FUNCTION_BLOCK FB_BECKHOFF_AxisController
(*

The function block used to control axis.

Constructor: 		Patryk Panylo
Company:		E. Riexinger GmbH
Date:			23.04.2015
Version:			1.00

Date:			Revision:		Who:				Comment
dd.mm.yyyy		x.xx			Initials			comment

*)
VAR_INPUT
	(* Input variables / Eingang Variablen *)
	bEnable						:BOOL;						(* Signal FB enable *)
	etMachineMode				:ET_MachineMode;			(* Machine mode *)
	etMachineState				:ET_MachineState;			(* Machine state *)
	bNoEStop					:BOOL;						(* No ermergency Stop / Keine Notaus *)
	bRegulatorOn				:BOOL;						(* Enable the power stage *)
	bReset						:BOOL;						(* Signal reset *)
	bCMDInterrupt				:BOOL;						(* Signal interrupt *)
	bTerminalOK					:BOOL;						(* Terminal Ok *)
	bExeReset					:BOOL;						(* Execute auto reset *)
	bExeSetPos					:BOOL;						(* Execute set position *)
	lrSetPosition				:LREAL;						(* Position value to which the axis position is to be set. *)
	bExeGearIn					:BOOL;						(* Execute gear in *)
	bExeGearOut					:BOOL;						(* Execute gear out *)
	dnRatioNumerator			:DINT;						(* Gear ratio numerator. Alternatively, the gear ratio can be specified in the numerator as a floating comma value, if the denominator is 1. *)
	udnRatioDenominator			:UDINT;						(* Gear ratio denominator *)
	lrOverride					:LREAL;						(* Override 100% percent *)
	bWithAbsoluteEncoder		:BOOL; 						(* Encoder is an absolute one / Absolutwertgeber *)
	bPosLagMonitoringEn			:BOOL;						(* Enable position lag monitoring *)
	lrPositionBias				:LREAL;						(* Position bias *)
	bHWSignalLimitMax			:BOOL;						(* Signal position limit switch maximum *)
	bHWSignalLimitMin			:BOOL;						(* Signal position limit switch minimum *)
	lrSoftLimitMax				:LREAL; 					(* Position limit switch maximum *)
	lrSoftLimitMin				:LREAL; 					(* Position limit switch minimum *)
	lrAcceleration				:LREAL;						(* Value of the acceleration (always positive) *)
	lrDeceleration				:LREAL;						(* Value of deceleration (always positive) *)
	lrJerk						:LREAL;						(* Value of jerk (always positive) *)
	lrActTemp					:LREAL;						(* Current temperatur *)
	tAdsTimeOut 				:TIME := T#2S;				(* Timout for ads commands *)
END_VAR
VAR_OUTPUT
	(* Output variables / Ausgang Variablen *)
	bStatus						:BOOL;						(* Feedback *)
	bStatusDelay				:BOOL;						(* Feedback delay *)
	bReseted					:BOOL;						(* Reset completed *)
	bError						:BOOL;						(* Controller error *)
	bErrorInit					:BOOL;						(* Controller initialization error *)
	udnErrorNo					:UDINT;						(* Error number *)
	lrActPos					:LREAL;						(* Actual position *)
	lrSetPos					:LREAL;						(* Set position *)
	lrActAbsPos					:LREAL;						(* Actual absolut position *)
	lrActVelo					:LREAL;						(* Actual velocity *)
	bNotMoving					:BOOL;						(* Status of moving *)
	bReferenced					:BOOL;						(* Referenced *)
	bCoupled					:BOOL;						(* Coupled *)
	lrVeloLimitMax				:LREAL;						(* Velocity limit maximum *)
	lrAccLimitMax				:LREAL;						(* Acceleration limit maximum *)
	lrDecLimitMax				:LREAL;						(* Deceleration limit maximum *)
	lrJerkLimitMax				:LREAL;						(* Jerk limit maximum *)
	bHardLimitMaxExceeded		:BOOL;						(* Position limit switch maximum is exceeded *)
	bHardLimitMinExceeded		:BOOL;						(* Position limit switch minimum is exceeded *)
	bSoftLimitMaxExceeded		:BOOL;						(* Position limit switch maximum is exceeded *)
	bSoftLimitMinExceeded		:BOOL;						(* Position limit switch minimum is exceeded *)
END_VAR
VAR_IN_OUT
	Axis						:AXIS_REF;					(* The AXIS_REF data type  is an interface between the PLC and the NC and contains axis information *)
	MasterAxis					:AXIS_REF;					(* The AXIS_REF data type  is an interface between the PLC and the NC and contains axis information *)
END_VAR
VAR
	(* Enummerations *)

	(* Variables *)
	etAxisGetLimits				:ET_BECKHOFF_AxisGetLimits;
	bGetLimitsExe				:BOOL;						(* Progam execute *)
	bGetLimitsDone 				:BOOL;                      (* Program done *)
	bGetLimitsBusy 				:BOOL;                      (* Program busy *)
	bGetLimitsError 			:BOOL;                      (* Program error *)
	bGetLimitsInitDone 			:BOOL;                      (* Program initialization done *)
	udnGetLimitsErrorNo 		:UDINT;                     (* Error number *)
	unGetValueWatchdog			:UINT;

	etAxisSetLimits				:ET_BECKHOFF_AxisSetLimits;
	bSetLimitsExe				:BOOL;						(* Progam execute *)
	bSetLimitsDone 				:BOOL;                      (* Program done *)
	bSetLimitsBusy 				:BOOL;                      (* Program busy *)
	bSetLimitsError 			:BOOL;                      (* Program error *)
	bSetLimitsInitDone 			:BOOL;                      (* Program initialization done *)
	bSetLimitsInitError 		:BOOL;                      (* Program initialization error *)
	udnSetLimitsErrorNo 		:UDINT;                     (* Error number *)
	unSetValueWatchdog			:UINT;

	tStatusDelay				:TIME := T#1S;				(* Status delay time *)
	tRegulatorOffDelay			:TIME := T#50MS;			(* Regulator off delay time *)

	dwReferenceSystem			:DWORD;						(* Reference system: 0 - INC, 1 - ABS, 2 - ABS MODULO *)
	lrPositionBiasCache			:LREAL;						(* Position bias *)
	lrSoftLimitMaxCache			:LREAL; 					(* Position limit switch maximum *)
	lrSoftLimitMinCache			:LREAL; 					(* Position limit switch minimum *)

	tonFirstInit				:TON;						(* First initialization *)
	bFirstTime					:BOOL;

	(* References *)

	(* Interfaces *)

	(* Instances *)
	fbMcPower					:MC_Power;					(* The function block is used to enable for an axis *)
	rtNoEStop					:R_TRIG;
	tofRegulatorOn				:TOF;						(* Delay controller disable *)
	tonStatusDelay				:TON;						(* Delay controller enabled status *)
	fbMcReset					:MC_Reset;					(* An axis reset is carried out with the function block *)
	fbMcSetPosition				:MC_SetPosition;			(* Sets the current axis position to a parameterisable value. *)
	fbMcGearIn					:MC_GearInDyn;				(* The function block is used to couples a slave axis to a master axis using a floating point gear ratio. *)
	fbMcGearOut					:MC_GearOut;				(* The function block  is used to decoupling the slave from the master axis.  *)
	fbMcReadParameter 			:MC_ReadParameter;			(* The function block is used to read an axis parameter. *)
	fbMcWriteParameter 			:MC_WriteParameter;			(* The function block is used to write an axis parameter. *)
	fbMcWriteBoolParameter 		:MC_WriteBoolParameter;		(* The function block is used to write bool value an axis parameter. *)
	fbAdsWrite					:ADSWRITE;					(* The function block permits execution of an ADS write command, for the transfer of data to an ADS device. *)
	fbAdsRead					:ADSREAD;					(* The function block permits execution of an ADS read command, for the transfer of data to an ADS device. *)
	tofRepeateSetLimitsInit		:TOF;
	tofRepeateGetLimitsInit		:TOF;
	tonCoupled					:TON;
END_VAR
VAR CONSTANT
	dwIdxGrMainPara				:DWORD := 16#00004000;		(* Index group for main parameters of axis *)
	dwIdxGrNCEncPara			:DWORD := 16#00005000;		(* Index group for nc-encoder parameters of axis *)
	dwIdxGrNCCtrlPara			:DWORD := 16#00006000;		(* Index group for nc-controller parameters of axis *)
	dwIdxGrNCDrivePara			:DWORD := 16#00007000;		(* Index group for nc-drive parameters of axis *)
	
	tFirstInit					:TIME := T#2S;				(* First initialization *)
	tRepeateInit				:TIME := T#1S;				(* Repeate initialization *)
	
	unWatchdogMax				:UINT := 150;
END_VAR

IF NOT bEnable							(* Signal FB enable *)
THEN
	bStatus := FALSE;						(* Feedback *)
	bStatusDelay := FALSE;				(* Feedback *)
	bError := FALSE;						(* Controller error *)
	udnErrorNo := 0;						(* Error number *)

	bFirstTime := FALSE;
	RETURN;
END_IF

IF NOT bFirstTime
THEN
	tonFirstInit(IN := FALSE);					(* Program execute *)
	bGetLimitsDone := FALSE;                                	(* Program done *)
	bGetLimitsBusy := FALSE;                                 	(* Program not busy *)
	bGetLimitsError := FALSE;                                 	(* Program not error *)
	bGetLimitsInitDone := FALSE;				(* Program initialization done *)
	udnGetLimitsErrorNo := 0;                                 		(* Error number *)
	unGetValueWatchdog := 0;

	etAxisGetLimits := ET_BECKHOFF_AxisGetLimits.eWaitExecute;       			(* Next step *)

	bSetLimitsExe := FALSE;					(* Program execute *)
	bSetLimitsDone := FALSE;                                	(* Program done *)
	bSetLimitsBusy := FALSE;                                 	(* Program not busy *)
	bSetLimitsError := FALSE;                                	 	(* Program not error *)
	bSetLimitsInitDone := FALSE;                            	(* Program initialization done *)
	bSetLimitsInitError := FALSE;				(* Program initialization error *)
	udnSetLimitsErrorNo := 0;                                 		(* Error number *)
	unSetValueWatchdog := 0;
	
	etAxisSetLimits := ET_BECKHOFF_AxisSetLimits.eWaitExecute;       			(* Next step *)

	(* Actual position *)
	lrActAbsPos := Axis.NcToPlc.ActPos;
	lrActAbsPos := F_LRealRound(lrReal := lrActAbsPos, usiPrecision := 3);

	bFirstTime := TRUE;
END_IF;

A_MCPower();
A_MCReset();
A_MCSetPosition();
A_MCGearCoupling();
A_Utility();
A_GetLimits();
A_SetLimits();
A_Error();

(* Actual position *)
lrActPos := Axis.NcToPlc.ActPos;
lrActPos := F_LRealRound(lrReal := lrActPos, usiPrecision := 2);

(* Set position *)
lrSetPos := Axis.NcToPlc.SetPos;
lrSetPos := F_LRealRound(lrReal := lrSetPos, usiPrecision := 2);

(* Actual velocity *)
lrActVelo := Axis.NcToPlc.ActVelo;
lrActVelo := F_LRealRound(lrReal := lrActVelo, usiPrecision := 2);

(* Current engine torque *)
(*nActEngineTorque := Axis.stNcToPlc.stCommandPositioning.nActEngineTorque;*)

(* Reference signal *)
bReferenced := Axis.NcToPlc.StateDWord.1;                               (* In Reference *)


(* Status not moving *)
bNotMoving := Axis.NcToPlc.StateDWord.2;

(* Status coupling *)
tonCoupled(
	IN := Axis.NcToPlc.CoupleState = 2
		  OR Axis.NcToPlc.CoupleState = 3,
	PT := T#200MS
);
bCoupled := tonCoupled.Q;

ACTION A_Error:

bError := fbMcPower.Error
		OR fbMcReset.Error
	  	OR fbMcSetPosition.Error
		OR fbMcGearIn.Error
		OR fbMcGearOut.Error
		OR Axis.NcToPlc.StateDWord.31
		OR MasterAxis.NcToPlc.StateDWord.31;

bErrorInit := bGetLimitsError
		      OR bSetLimitsError;
END_ACTION

ACTION A_GetLimits:

(* Status hardware limit switch *)
bHardLimitMaxExceeded := bHWSignalLimitMax;						(* Position limit switch maximum is exceeded *)
bHardLimitMinExceeded := bHWSignalLimitMin;						(* Position limit switch minimum is exceeded *)

(* Status software limit switch *)
bSoftLimitMaxExceeded := Axis.NcToPlc.StateDWord.27 AND lrSoftLimitMax <> lrSoftLimitMin;	(* Position limit switch maximum is exceeded *)
bSoftLimitMinExceeded := Axis.NcToPlc.StateDWord.26 AND lrSoftLimitMax <> lrSoftLimitMin;		(* Position limit switch minimum is exceeded *)

(* Get limits execute *)
tofRepeateGetLimitsInit(
	IN := bGetLimitsError,
	PT := tRepeateInit
);

tonFirstInit(
	IN:= bTerminalOK
		 AND NOT bGetLimitsInitDone,
	PT := tFirstInit
);

bGetLimitsExe := (tonFirstInit.Q
				  OR bGetLimitsInitDone)
				  AND NOT tofRepeateGetLimitsInit.Q;

(* Get axis limits *)
CASE etAxisGetLimits OF

	ET_BECKHOFF_AxisGetLimits.eWaitExecute:
		IF bGetLimitsExe
		   AND bTerminalOK
		THEN
			unGetValueWatchdog := 0;
			bGetLimitsDone := FALSE;                                	(* Program done *)
			bGetLimitsBusy := FALSE;                                 	(* Program not busy *)
			bGetLimitsError := FALSE;                                 	(* Program not error *)
			udnGetLimitsErrorNo := 0;                                 	(* Error number *)

			fbMcReadParameter(
				Enable:= FALSE,
				ReadMode := READMODE_ONCE,
				Axis := Axis
			);

			fbAdsRead(
				NETID := '',
				READ := FALSE,
				TMOUT := tAdsTimeOut
			);
			
			etAxisGetLimits := ET_BECKHOFF_AxisGetLimits.eReadVeloMax;         		(* Next step *)
		END_IF

	ET_BECKHOFF_AxisGetLimits.eReadVeloMax:
		fbMcReadParameter.Enable := TRUE;
		fbMcReadParameter.ParameterNumber:= MaxVelocityAppl;

		unGetValueWatchdog := unGetValueWatchdog + 1;
		
		IF fbMcReadParameter.Busy
		THEN
			etAxisGetLimits := ET_BECKHOFF_AxisGetLimits.eWfReadVeloMax;         		(* Next step *)

		ELSIF fbMcReadParameter.Error
		THEN
			fbMcReadParameter(
				Enable:= FALSE,
				Axis := Axis
			);

			udnGetLimitsErrorNo := 1;                                 	(* Error number *)
			
			etAxisGetLimits := ET_BECKHOFF_AxisGetLimits.eError;         		(* Next step *)

		END_IF

	ET_BECKHOFF_AxisGetLimits.eWfReadVeloMax:
		IF NOT fbMcReadParameter.Busy
		     AND NOT fbMcReadParameter.Error
		THEN
			fbMcReadParameter(
				Enable:= FALSE,
				Axis := Axis
			);

			lrVeloLimitMax := fbMcReadParameter.Value;

			unGetValueWatchdog := 0;
			
			etAxisGetLimits := ET_BECKHOFF_AxisGetLimits.eReadAccMax;         		(* Next step *)

		ELSIF fbMcReadParameter.Error
		THEN
			fbMcReadParameter(
				Enable:= FALSE,
				Axis := Axis
			);

			udnGetLimitsErrorNo := 2;                                 	(* Error number *)
			
			etAxisGetLimits := ET_BECKHOFF_AxisGetLimits.eError;         		(* Next step *)

		END_IF

	ET_BECKHOFF_AxisGetLimits.eReadAccMax:
		fbMcReadParameter.Enable := TRUE;
		fbMcReadParameter.ParameterNumber:= MaxAccelerationAppl;

		unGetValueWatchdog := unGetValueWatchdog + 1;
		
		IF fbMcReadParameter.Busy
		THEN
			etAxisGetLimits := ET_BECKHOFF_AxisGetLimits.eWfReadAccMax;         		(* Next step *)

		ELSIF fbMcReadParameter.Error
		THEN
			fbMcReadParameter(
				Enable:= FALSE,
				Axis := Axis
			);

			udnGetLimitsErrorNo := 3;                                 	(* Error number *)
			
			etAxisGetLimits := ET_BECKHOFF_AxisGetLimits.eError;         		(* Next step *)

		END_IF

	ET_BECKHOFF_AxisGetLimits.eWfReadAccMax:
		IF NOT fbMcReadParameter.Busy
		     AND NOT fbMcReadParameter.Error
		THEN
			fbMcReadParameter(
				Enable:= FALSE,
				Axis := Axis
			);

			lrAccLimitMax := fbMcReadParameter.Value;

			unGetValueWatchdog := 0;
			
			etAxisGetLimits := ET_BECKHOFF_AxisGetLimits.eReadDecMax;         		(* Next step *)

		ELSIF fbMcReadParameter.Error
		THEN
			fbMcReadParameter(
				Enable:= FALSE,
				Axis := Axis
			);

			udnGetLimitsErrorNo := 4;                                 	(* Error number *)
			
			etAxisGetLimits := ET_BECKHOFF_AxisGetLimits.eError;         		(* Next step *)

		END_IF

	ET_BECKHOFF_AxisGetLimits.eReadDecMax:
		fbMcReadParameter.Enable := TRUE;
		fbMcReadParameter.ParameterNumber:= MaxDecelerationAppl;

		unGetValueWatchdog := unGetValueWatchdog + 1;
		
		IF fbMcReadParameter.Busy
		THEN
			etAxisGetLimits := ET_BECKHOFF_AxisGetLimits.eWfReadDecMax;         		(* Next step *)

		ELSIF fbMcReadParameter.Error
		THEN
			fbMcReadParameter(
				Enable:= FALSE,
				Axis := Axis
			);

			udnGetLimitsErrorNo := 5;                                 	(* Error number *)
			
			etAxisGetLimits := ET_BECKHOFF_AxisGetLimits.eError;         		(* Next step *)

		END_IF

	ET_BECKHOFF_AxisGetLimits.eWfReadDecMax:
		IF NOT fbMcReadParameter.Busy
		     AND NOT fbMcReadParameter.Error
		THEN
			fbMcReadParameter(
				Enable:= FALSE,
				Axis := Axis
			);

			lrDecLimitMax := fbMcReadParameter.Value;

			unGetValueWatchdog := 0;
			
			etAxisGetLimits := ET_BECKHOFF_AxisGetLimits.eReadJerkMax;         		(* Next step *)

		ELSIF fbMcReadParameter.Error
		THEN
			fbMcReadParameter(
				Enable:= FALSE,
				Axis := Axis
			);

			udnGetLimitsErrorNo := 6;                                 	(* Error number *)
			
			etAxisGetLimits := ET_BECKHOFF_AxisGetLimits.eError;         		(* Next step *)

		END_IF

	ET_BECKHOFF_AxisGetLimits.eReadJerkMax:
		fbMcReadParameter.Enable := TRUE;
		fbMcReadParameter.ParameterNumber:= MaxJerkAppl;

		unGetValueWatchdog := unGetValueWatchdog + 1;
		
		IF fbMcReadParameter.Busy
		THEN
			etAxisGetLimits := ET_BECKHOFF_AxisGetLimits.eWfReadJerkMax;         		(* Next step *)

		ELSIF fbMcReadParameter.Error
		THEN
			fbMcReadParameter(
				Enable:= FALSE,
				Axis := Axis
			);

			udnGetLimitsErrorNo := 7;                                 	(* Error number *)
			
			etAxisGetLimits := ET_BECKHOFF_AxisGetLimits.eError;         		(* Next step *)

		END_IF

	ET_BECKHOFF_AxisGetLimits.eWfReadJerkMax:
		IF NOT fbMcReadParameter.Busy
		     AND NOT fbMcReadParameter.Error
		THEN
			fbMcReadParameter(
				Enable:= FALSE,
				Axis := Axis
			);

			lrJerkLimitMax := fbMcReadParameter.Value;

			unGetValueWatchdog := 0;
			
			etAxisGetLimits := ET_BECKHOFF_AxisGetLimits.eReadSoftLimitMax;         		(* Next step *)

		ELSIF fbMcReadParameter.Error
		THEN
			fbMcReadParameter(
				Enable:= FALSE,
				Axis := Axis
			);

			udnGetLimitsErrorNo := 8;                                 	(* Error number *)
			
			etAxisGetLimits := ET_BECKHOFF_AxisGetLimits.eError;         		(* Next step *)

		END_IF

	ET_BECKHOFF_AxisGetLimits.eReadSoftLimitMax:
		fbMcReadParameter.Enable := TRUE;
		fbMcReadParameter.ParameterNumber:= SWLimitPos;

		unGetValueWatchdog := unGetValueWatchdog + 1;
		
		IF fbMcReadParameter.Busy
		THEN
			etAxisGetLimits := ET_BECKHOFF_AxisGetLimits.eWfReadSoftLimitMax;         		(* Next step *)

		ELSIF fbMcReadParameter.Error
		THEN
			fbMcReadParameter(
				Enable:= FALSE,
				Axis := Axis
			);

			udnGetLimitsErrorNo := 9;                                 	(* Error number *)
			
			etAxisGetLimits := ET_BECKHOFF_AxisGetLimits.eError;         		(* Next step *)

		END_IF

	ET_BECKHOFF_AxisGetLimits.eWfReadSoftLimitMax:
		IF NOT fbMcReadParameter.Busy
		     AND NOT fbMcReadParameter.Error
		THEN
			fbMcReadParameter(
				Enable:= FALSE,
				Axis := Axis
			);

			lrSoftLimitMax := fbMcReadParameter.Value;

			unGetValueWatchdog := 0;
			
			etAxisGetLimits := ET_BECKHOFF_AxisGetLimits.eReadSoftLimitMin;         		(* Next step *)

		ELSIF fbMcReadParameter.Error
		THEN
			fbMcReadParameter(
				Enable:= FALSE,
				Axis := Axis
			);

			udnGetLimitsErrorNo := 10;                                 	(* Error number *)
			
			etAxisGetLimits := ET_BECKHOFF_AxisGetLimits.eError;         		(* Next step *)

		END_IF

	ET_BECKHOFF_AxisGetLimits.eReadSoftLimitMin:
		fbMcReadParameter.Enable := TRUE;
		fbMcReadParameter.ParameterNumber:= SWLimitNeg;

		unGetValueWatchdog := unGetValueWatchdog + 1;
		
		IF fbMcReadParameter.Busy
		THEN
			etAxisGetLimits := ET_BECKHOFF_AxisGetLimits.eWfReadSoftLimitMin;         		(* Next step *)

		ELSIF fbMcReadParameter.Error
		THEN
			fbMcReadParameter(
				Enable:= FALSE,
				Axis := Axis
			);

			udnGetLimitsErrorNo := 11;                                 	(* Error number *)
			
			etAxisGetLimits := ET_BECKHOFF_AxisGetLimits.eError;         		(* Next step *)

		END_IF

	ET_BECKHOFF_AxisGetLimits.eWfReadSoftLimitMin:
		IF NOT fbMcReadParameter.Busy
		     AND NOT fbMcReadParameter.Error
		THEN
			fbMcReadParameter(
				Enable:= FALSE,
				Axis := Axis
			);

			lrSoftLimitMin := fbMcReadParameter.Value;

			unGetValueWatchdog := 0;
			
			etAxisGetLimits := ET_BECKHOFF_AxisGetLimits.eDone;         		(* Next step *)

		ELSIF fbMcReadParameter.Error
		THEN
			fbMcReadParameter(
				Enable:= FALSE,
				Axis := Axis
			);

			udnGetLimitsErrorNo := 12;                                 	(* Error number *)
			
			etAxisGetLimits := ET_BECKHOFF_AxisGetLimits.eError;         		(* Next step *)

		END_IF
	
	ET_BECKHOFF_AxisGetLimits.eDone:
		bGetLimitsDone := TRUE;                                     		(* Program done, in position *)
		bGetLimitsBusy := FALSE;                                     		(* Program not busy *)
		bGetLimitsInitDone := TRUE;                             		(* Program initialization done *)

		etAxisGetLimits := ET_BECKHOFF_AxisGetLimits.eNoExecute;            	(* Next step *)

	ET_BECKHOFF_AxisGetLimits.eError:
		bGetLimitsDone := FALSE;                                     		(* Program done, in position *)
		bGetLimitsError := TRUE;                                     		(* Program error *)
		bGetLimitsBusy := FALSE;                                     		(* Program not busy *)
		bGetLimitsInitDone := FALSE;                             		(* Program initialization done *)

		etAxisGetLimits := ET_BECKHOFF_AxisGetLimits.eNoExecute;           	(* Next step *)

	ET_BECKHOFF_AxisGetLimits.eNoExecute:
		IF NOT bGetLimitsExe
		THEN
			bGetLimitsDone := FALSE;                                     		(* Program done, in position *)
			bGetLimitsError := FALSE;                                     		(* Program error *)
			bGetLimitsBusy := FALSE;                                     		(* Program not busy *)

			etAxisGetLimits := ET_BECKHOFF_AxisGetLimits.eWaitExecute;       (* Next step *)
		END_IF

END_CASE;

fbMcReadParameter(
	ReadMode := READMODE_ONCE,
	Axis := Axis
);
END_ACTION

ACTION A_MCGearCoupling:

(* The function block MC_GearInDyn couples a slave axis to a master axis using a floating point gear ratio. The gear ratio can be dynamically modified every PLC cycle as long as the Execute input is TRUE *)
IF udnRatioDenominator = 0
THEN
	fbMCGearIn.GearRatio := 0;
ELSE
	fbMCGearIn.GearRatio:= dnRatioNumerator / udnRatioDenominator;
END_IF


IF NOT bCMDInterrupt
THEN

	(* The function block MC_GearIn used to coupling with ratio between the velocity of the slave and master axis  *)
	fbMCGearIn(
		Enable := bExeGearIn,
		Acceleration := lrAcceleration,
		Deceleration := lrDeceleration,
		Jerk := lrJerk,
		Options := ,
		Master := MasterAxis,
		Slave := Axis
	);
	
	(* The function block MC_GearOut used to decoupling the Slave from the Master axis.  *)
	fbMCGearOut(
		Execute := bExeGearOut,
		Slave := Axis,
	);

	(* Weiter für die GearIn und GearOut entwickeln*)
	(*Axis.bCmdInterrupted := FALSE;*)

ELSE
	(* The function block MC_GearIn used to coupling with ratio between the velocity of the slave and master axis  *)
	fbMCGearIn(
		Enable := FALSE,
		Master := MasterAxis,
		Slave := Axis
	);

	(* The function block MC_GearOut used to decoupling the Slave from the Master axis.  *)
	fbMCGearOut(
		Execute := FALSE,
		Slave := Axis
	);

	(*Axis.bCmdInterrupted := TRUE;*)
END_IF
END_ACTION

ACTION A_MCPower:

tofRegulatorOn(
	IN := bRegulatorOn,
	PT := tRegulatorOffDelay
);

fbMCPower(
	Enable := tofRegulatorOn.Q
			OR Axis.Status.Moving,
	Enable_Positive := (bRegulatorOn
					AND NOT bHWSignalLimitMax)                          			(* HW limit switch maximum *)
					OR Axis.NcToPlc.HomingState <> 0,
	Enable_Negative := (bRegulatorOn
					   AND NOT bHWSignalLimitMin)                         			(* HW Limit switch minimum *)
					   OR Axis.NcToPlc.HomingState <> 0,
	Override := LIMIT(0.0, lrOverride, 100.0),
	Axis := Axis,
	Status => bStatus,
);

tonStatusDelay(
	IN := fbMCPower.Status,
	PT := SEL(etMachineMode = ET_MachineMode_eManual, tStatusDelay, t#0s),
	Q => bStatusDelay
);
END_ACTION

ACTION A_MCReset:

rtNoEStop(CLK := bNoEStop);

fbMCReset(
	Execute := rtNoEStop.Q
			   OR (bReset
			   		AND Axis.NcToPlc.StateDWord.31)
			   OR bExeReset,
	Axis := Axis,
	Done => bReseted
 );
END_ACTION

ACTION A_MCSetPosition:

fbMCSetPosition(
	Execute := bExeSetPos,
	Position := SEL(lrSoftLimitMin <> lrSoftLimitMax, lrSetPosition, LIMIT(lrSoftLimitMin, lrSetPosition, lrSoftLimitMax)),
	Mode := FALSE,
	Options := ,
	Axis := Axis
);
END_ACTION

ACTION A_SetLimits:

(* Set limits execute *)
tofRepeateSetLimitsInit(
	IN := bSetLimitsError,
	PT := tRepeateInit
);

bSetLimitsExe := SEL(
						bSetLimitsInitDone,
						NOT bSetLimitsInitError,
						NOT bSetLimitsInitError
						AND (lrPositionBias <> lrPositionBiasCache
							   OR lrSoftLimitMaxCache <> lrSoftLimitMax
							   OR lrSoftLimitMinCache <> lrSoftLimitMin)
					);

(* Set axis limits *)
CASE etAxisSetLimits OF

	ET_BECKHOFF_AxisSetLimits.eWaitExecute:
		IF bSetLimitsExe
		   AND bTerminalOK
		   AND bNotMoving
		   AND bGetLimitsDone
		THEN
			unSetValueWatchdog := 0;
			bSetLimitsDone := FALSE;                                	(* Program done *)
			bSetLimitsBusy := FALSE;                                 	(* Program not busy *)
			bSetLimitsError := FALSE;                                	 	(* Program not error *)
			udnSetLimitsErrorNo := 0;                                 		(* Error number *)

			fbMcWriteParameter(
				Execute := FALSE,
				Axis := Axis
			);
	
			fbMcWriteBoolParameter(
				Execute := FALSE,
				Axis := Axis
			);
	
			fbAdsWrite(
				NETID := '',
				WRITE := FALSE,
				TMOUT := tAdsTimeOut
			 );

			etAxisSetLimits := ET_BECKHOFF_AxisSetLimits.eSetReferenceSystem;         		(* Next step *)

		END_IF;

	ET_BECKHOFF_AxisSetLimits.eSetReferenceSystem:
		dwReferenceSystem := BOOL_TO_DWORD(bWithAbsoluteEncoder);

		fbAdsWrite.PORT := 501;
		fbAdsWrite.WRITE := TRUE;
		fbAdsWrite.IDXGRP := dwIdxGrNCEncPara + Axis.NcToPlc.AxisId;
		fbAdsWrite.IDXOFFS := 16#00000019;
		fbAdsWrite.LEN := SIZEOF(dwReferenceSystem);
		fbAdsWrite.SRCADDR := ADR(dwReferenceSystem);

		unSetValueWatchdog := unSetValueWatchdog + 1;
		
		IF fbAdsWrite.Busy
		THEN
			etAxisSetLimits := ET_BECKHOFF_AxisSetLimits.eWfSetReferenceSystem;         		(* Next step *)

		ELSIF fbAdsWrite.ERR
		THEN
			fbAdsWrite(
				WRITE := FALSE,
			);

			udnSetLimitsErrorNo := 1;                                 		(* Error number *)
			
			etAxisSetLimits := ET_BECKHOFF_AxisSetLimits.eError;         		(* Next step *)

		END_IF

	ET_BECKHOFF_AxisSetLimits.eWfSetReferenceSystem:
		IF NOT fbAdsWrite.Busy
		     AND NOT fbAdsWrite.ERR
		THEN
			fbAdsWrite(
				WRITE := FALSE,
			);

			unSetValueWatchdog := 0;
			
			etAxisSetLimits := ET_BECKHOFF_AxisSetLimits.eSetPositionBias;         		(* Next step *)

		ELSIF fbAdsWrite.ERR
		THEN
			fbAdsWrite(
				WRITE := FALSE,
			);

			udnSetLimitsErrorNo := 2;                                 		(* Error number *)
			
			etAxisSetLimits := ET_BECKHOFF_AxisSetLimits.eError;         		(* Next step *)

		END_IF

	ET_BECKHOFF_AxisSetLimits.eSetPositionBias:
		IF bWithAbsoluteEncoder
		THEN
			lrPositionBiasCache := lrPositionBias;

			fbAdsWrite.PORT := 501;
			fbAdsWrite.WRITE := TRUE;
			fbAdsWrite.IDXGRP := dwIdxGrNCEncPara + Axis.NcToPlc.AxisId;
			fbAdsWrite.IDXOFFS := 16#00000007;
			fbAdsWrite.LEN := SIZEOF(lrPositionBiasCache);
			fbAdsWrite.SRCADDR := ADR(lrPositionBiasCache);
	
			unSetValueWatchdog := unSetValueWatchdog + 1;
			
			IF fbAdsWrite.Busy
			THEN
				etAxisSetLimits := ET_BECKHOFF_AxisSetLimits.eWfSetPositionBias;         		(* Next step *)
	
			ELSIF fbAdsWrite.ERR
			THEN
				fbAdsWrite(
					WRITE := FALSE,
				);
	
				udnSetLimitsErrorNo := 3;                                 		(* Error number *)
				
				etAxisSetLimits := ET_BECKHOFF_AxisSetLimits.eError;         		(* Next step *)
	
			END_IF
		ELSE
			etAxisSetLimits := ET_BECKHOFF_AxisSetLimits.eSetLimitPos;         		(* Next step *)

		END_IF

	ET_BECKHOFF_AxisSetLimits.eWfSetPositionBias:
		IF NOT fbAdsWrite.Busy
		     AND NOT fbAdsWrite.ERR
		THEN
			fbAdsWrite(
				WRITE := FALSE,
			);

			unSetValueWatchdog := 0;
			
			etAxisSetLimits := ET_BECKHOFF_AxisSetLimits.eSetLimitPos;         		(* Next step *)

		ELSIF fbAdsWrite.ERR
		THEN
			fbAdsWrite(
				WRITE := FALSE,
			);

			udnSetLimitsErrorNo := 4;                                 		(* Error number *)
			
			etAxisSetLimits := ET_BECKHOFF_AxisSetLimits.eError;         		(* Next step *)

		END_IF

	ET_BECKHOFF_AxisSetLimits.eSetLimitPos:
		lrSoftLimitMaxCache := lrSoftLimitMax;

		fbMcWriteParameter.Execute := TRUE;
		fbMcWriteParameter.ParameterNumber := SWLimitPos;
		fbMcWriteParameter.Value := lrSoftLimitMax;

		unSetValueWatchdog := unSetValueWatchdog + 1;
		
		IF fbMcWriteParameter.Busy
		THEN
			etAxisSetLimits := ET_BECKHOFF_AxisSetLimits.eWfSetLimitPos;         		(* Next step *)

		ELSIF fbMcWriteParameter.Error
		THEN
			fbMcWriteParameter(
				Execute := FALSE,
				Axis := Axis
			);

			udnSetLimitsErrorNo := 4;                                 		(* Error number *)
			
			etAxisSetLimits := ET_BECKHOFF_AxisSetLimits.eError;         		(* Next step *)

		END_IF

	ET_BECKHOFF_AxisSetLimits.eWfSetLimitPos:
		IF NOT fbMcWriteParameter.Busy
		     AND NOT fbMcWriteParameter.Error
		THEN
			fbMcWriteParameter(
				Execute := FALSE,
				Axis := Axis
			);

			unSetValueWatchdog := 0;
			
			etAxisSetLimits := ET_BECKHOFF_AxisSetLimits.eSetLimitNeg;         		(* Next step *)

		ELSIF fbMcWriteParameter.Error
		THEN
			fbMcWriteParameter(
				Execute := FALSE,
				Axis := Axis
			);

			udnSetLimitsErrorNo := 5;                                 		(* Error number *)
			
			etAxisSetLimits := ET_BECKHOFF_AxisSetLimits.eError;         		(* Next step *)

		END_IF

	ET_BECKHOFF_AxisSetLimits.eSetLimitNeg:
		lrSoftLimitMinCache := lrSoftLimitMin;

		fbMcWriteParameter.Execute := TRUE;
		fbMcWriteParameter.ParameterNumber := SWLimitNeg;
		fbMcWriteParameter.Value := lrSoftLimitMin;

		unSetValueWatchdog := unSetValueWatchdog + 1;
		
		IF fbMcWriteParameter.Busy
		THEN
			etAxisSetLimits := ET_BECKHOFF_AxisSetLimits.eWfSetLimitNeg;         		(* Next step *)

		ELSIF fbMcWriteParameter.Error
		THEN
			fbMcWriteParameter(
				Execute := FALSE,
				Axis := Axis
			);

			udnSetLimitsErrorNo := 6;                                 		(* Error number *)
			
			etAxisSetLimits := ET_BECKHOFF_AxisSetLimits.eError;         		(* Next step *)

		END_IF

	ET_BECKHOFF_AxisSetLimits.eWfSetLimitNeg:
		IF NOT fbMcWriteParameter.Busy
		     AND NOT fbMcWriteParameter.Error
		THEN
			fbMcWriteParameter(
				Execute := FALSE,
				Axis := Axis
			);

			unSetValueWatchdog := 0;
			
			etAxisSetLimits := ET_BECKHOFF_AxisSetLimits.eEnableLimitPos;         		(* Next step *)

		ELSIF fbMcWriteParameter.Error
		THEN
			fbMcWriteParameter(
				Execute := FALSE,
				Axis := Axis
			);

			udnSetLimitsErrorNo := 6;                                 		(* Error number *)
			
			etAxisSetLimits := ET_BECKHOFF_AxisSetLimits.eError;         		(* Next step *)

		END_IF

	ET_BECKHOFF_AxisSetLimits.eEnableLimitPos:
		fbMcWriteBoolParameter.Execute := TRUE;
		fbMcWriteBoolParameter.ParameterNumber := EnableLimitPos;
		fbMcWriteBoolParameter.Value := lrSoftLimitMax <> lrSoftLimitMin;

		unSetValueWatchdog := unSetValueWatchdog + 1;
		
		IF fbMcWriteBoolParameter.Busy
		THEN
			etAxisSetLimits := ET_BECKHOFF_AxisSetLimits.eWfEnableLimitPos;         		(* Next step *)

		ELSIF fbMcWriteBoolParameter.Error
		THEN
			fbMcWriteBoolParameter(
				Execute := FALSE,
				Axis := Axis
			);

			udnSetLimitsErrorNo := 7;                                 		(* Error number *)
			
			etAxisSetLimits := ET_BECKHOFF_AxisSetLimits.eError;         		(* Next step *)

		END_IF

	ET_BECKHOFF_AxisSetLimits.eWfEnableLimitPos:
		IF NOT fbMcWriteBoolParameter.Busy
		     AND NOT fbMcWriteBoolParameter.Error
		THEN
			fbMcWriteBoolParameter(
				Execute := FALSE,
				Axis := Axis
			);

			unSetValueWatchdog := 0;
			
			etAxisSetLimits := ET_BECKHOFF_AxisSetLimits.eEnableLimitNeg;         		(* Next step *)

		ELSIF fbMcWriteBoolParameter.Error
		THEN
			fbMcWriteBoolParameter(
				Execute := FALSE,
				Axis := Axis
			);

			udnSetLimitsErrorNo := 8;                                 		(* Error number *)
			
			etAxisSetLimits := ET_BECKHOFF_AxisSetLimits.eError;         		(* Next step *)

		END_IF

	ET_BECKHOFF_AxisSetLimits.eEnableLimitNeg:
		fbMcWriteBoolParameter.Execute := TRUE;
		fbMcWriteBoolParameter.ParameterNumber := EnableLimitNeg;
		fbMcWriteBoolParameter.Value := lrSoftLimitMax <> lrSoftLimitMin;

		unSetValueWatchdog := unSetValueWatchdog + 1;
		
		IF fbMcWriteBoolParameter.Busy
		THEN
			etAxisSetLimits := ET_BECKHOFF_AxisSetLimits.eWfEnableLimitNeg;         		(* Next step *)

		ELSIF fbMcWriteBoolParameter.Error
		THEN
			fbMcWriteBoolParameter(
				Execute := FALSE,
				Axis := Axis
			);

			udnSetLimitsErrorNo := 9;                                 		(* Error number *)
			
			etAxisSetLimits := ET_BECKHOFF_AxisSetLimits.eError;         		(* Next step *)

		END_IF

	ET_BECKHOFF_AxisSetLimits.eWfEnableLimitNeg:
		IF NOT fbMcWriteBoolParameter.Busy
		     AND NOT fbMcWriteBoolParameter.Error
		THEN
			fbMcWriteBoolParameter(
				Execute := FALSE,
				Axis := Axis
			);

			unSetValueWatchdog := 0;
			
			etAxisSetLimits := ET_BECKHOFF_AxisSetLimits.eEnablePosLagMonitoring;         		(* Next step *)

		ELSIF fbMcWriteBoolParameter.Error
		THEN
			fbMcWriteBoolParameter(
				Execute := FALSE,
				Axis := Axis
			);

			udnSetLimitsErrorNo := 10;                                 		(* Error number *)
			
			etAxisSetLimits := ET_BECKHOFF_AxisSetLimits.eError;         		(* Next step *)

		END_IF

	ET_BECKHOFF_AxisSetLimits.eEnablePosLagMonitoring:
		fbMcWriteBoolParameter.Execute := TRUE;
		fbMcWriteBoolParameter.ParameterNumber := EnablePosLagMonitoring;
		fbMcWriteBoolParameter.Value := bPosLagMonitoringEn;

		unSetValueWatchdog := unSetValueWatchdog + 1;
		
		IF fbMcWriteBoolParameter.Busy
		THEN
			etAxisSetLimits := ET_BECKHOFF_AxisSetLimits.eWfEnablePosLagMonitoring;         		(* Next step *)

		ELSIF fbMcWriteBoolParameter.Error
		THEN
			fbMcWriteBoolParameter(
				Execute := FALSE,
				Axis := Axis
			);

			udnSetLimitsErrorNo := 11;                                 		(* Error number *)
			
			etAxisSetLimits := ET_BECKHOFF_AxisSetLimits.eError;         		(* Next step *)

		END_IF

	ET_BECKHOFF_AxisSetLimits.eWfEnablePosLagMonitoring:
		IF NOT fbMcWriteBoolParameter.Busy
		     AND NOT fbMcWriteBoolParameter.Error
		THEN
			fbMcWriteBoolParameter(
				Execute := FALSE,
				Axis := Axis
			);

			unSetValueWatchdog := 0;
			
			etAxisSetLimits := ET_BECKHOFF_AxisSetLimits.eDone;         		(* Next step *)

		ELSIF fbMcWriteBoolParameter.Error
		THEN
			fbMcWriteBoolParameter(
				Execute := FALSE,
				Axis := Axis
			);

			udnSetLimitsErrorNo := 12;                                 		(* Error number *)
			
			etAxisSetLimits := ET_BECKHOFF_AxisSetLimits.eError;         		(* Next step *)

		END_IF

	ET_BECKHOFF_AxisSetLimits.eDone:
		bSetLimitsDone := TRUE;                                     		(* Program done, in position *)
		bSetLimitsBusy := FALSE;                                     		(* Program not busy *)
		bSetLimitsInitDone := TRUE;                             		(* Program initialization done *)

		etAxisSetLimits := ET_BECKHOFF_AxisSetLimits.eNoExecute;            	(* Next step *)

	ET_BECKHOFF_AxisSetLimits.eError:
		bSetLimitsDone := FALSE;                                     		(* Program done, in position *)
		bSetLimitsError := TRUE;                                     		(* Program error *)
		bSetLimitsBusy := FALSE;                                     		(* Program not busy *)
		bSetLimitsInitDone := FALSE;                             		(* Program initialization done *)

		etAxisSetLimits := ET_BECKHOFF_AxisSetLimits.eNoExecute;           	(* Next step *)

	ET_BECKHOFF_AxisSetLimits.eNoExecute:
		IF NOT bSetLimitsExe
		THEN
			bSetLimitsDone := FALSE;                                     		(* Program done, in position *)
			bSetLimitsError := FALSE;                                     		(* Program error *)
			bSetLimitsBusy := FALSE;                                     		(* Program not busy *)

			etAxisSetLimits := ET_BECKHOFF_AxisSetLimits.eWaitExecute;       (* Next step *)
		END_IF;

END_CASE;

fbMcWriteParameter(
	Axis := Axis
);

fbMcWriteBoolParameter(
	Axis := Axis
);

fbAdsWrite(
	NETID := '',
	TMOUT := tAdsTimeOut
 );
END_ACTION

ACTION A_Utility:

;
END_ACTION

END_FUNCTION_BLOCK

(* stored: Version 1.1.0.1, ProductVersion 3.1.4024.15
   POU FB_BECKHOFF_AxisController: Id {a7ff8751-94dc-481c-9120-4c27038cb85f}, SpecialFunc None
   Action A_Error: Id {020e17fe-7030-4d31-aed3-afb70cfda31a}
   Action A_GetLimits: Id {db11ab12-1104-4117-af2e-a8d657fbdea2}
   Action A_MCGearCoupling: Id {e1ffcbd7-7345-4d77-a0e0-64700b5e2332}
   Action A_MCPower: Id {e0593327-f1c0-42de-b721-674d8122d312}
   Action A_MCReset: Id {691769cd-5519-4703-92bf-05a64d07e631}
   Action A_MCSetPosition: Id {8ceb89c6-b87a-452d-9f5b-0d686dd7adcd}
   Action A_SetLimits: Id {fb969af6-e3df-41c1-ad19-f006e25f456a}
   Action A_Utility: Id {a98b9573-80c9-47c2-b6dd-ff37a945cd50} *)
